// TIA Portal V20 export
// export: Created 2025-07-07T08:55:10.1278921Z, ExportSetting None, DisplayName Totally Integrated Automation Portal, DisplayVersion V20 Update 5, DisplayName TIA Portal Openness, DisplayVersion V20 Update 5, DisplayName TIA Portal Version Control Interface, DisplayVersion V20, DisplayName SINAMICS Startdrive Advanced, DisplayVersion V20, DisplayName SINAMICS Startdrive G130, G150, S120, S150, SINAMICS MV, S210, DisplayVersion V20, DisplayName SINAMICS Startdrive G110M, G120, G120C, G120D, G120P, G115D, DisplayVersion V20, DisplayName STEP 7 Professional, DisplayVersion V20 Update 5, DisplayName STEP 7 Safety, DisplayVersion V20, DisplayName WinCC Advanced, DisplayVersion V20 Update 5
DATA_BLOCK "FB_PR_CentreStand_Fix_Seq_V12_V14_DB"   // DB1
// stored: InstanceOfName FB_PR_CentreStand_Fix_Seq_V12_V14, InstanceOfType FB
"FB_PR_CentreStand_Fix_Seq_V12_V14"
   // VAR_INPUT
   //    iAutoRunning : Bool;
   //    iFixClamp : Bool;
   //    iFixEmpty : Bool;
   //    iFixTrayPresent : Bool;
   //    iFixUnclamp : Bool;
   //    iR1DropOver : Bool;
   //    iR1PickOver : Bool;
   //    iR2OperationOver : Bool;
   //    iR2ServiceActivated : Bool;
   //    iReset_fault : Bool;
   //    iRobotOutofZone : Bool;
   //    iSstMode : Bool;
   //    iSstPB : Bool;
   // END_VAR
   // VAR_OUTPUT
   //    qFixClamp : Bool;
   //    qFixUnclamp : Bool;
   //    qR1ReadytoDropTray : Bool;
   //    qR1ReadytoPickTray : Bool;
   //    qR2OperationStart : Bool;
   // END_VAR
   // VAR_IN_OUT
   //    iqR2ServiceActive : Bool;
   //    iqR2ServiceCompleted : Bool;
   // END_VAR
BEGIN
END_DATA_BLOCK
